{attribute 'qualified_only'}
{attribute 'strict'}
{attribute 'to_string'}
TYPE E_StatusIndicator :
(
    Init := 10,
    Wait := 11,
    Complete := 12,
    Closed := 13,
    Opened := 14,
    Done := 15,
    // Special states
    HardReset := 80,
    SoftReset := 81
);
END_TYPE

(* stored: Version 1.1.0.1
   DUT E_StatusIndicator: Id {b89278ed-6a01-4923-a697-63d6bcfefc4c} *)
